FUNCTION_BLOCK CASCADE_CONTROL (* Migrated from IEC 61131-3 ST *)
  (* Standard: 61499-2 *)
  (* Version 1.0, 2026-11-06, st2fb *)
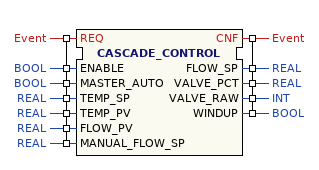
  EVENT_INPUT
    REQ WITH ENABLE, MASTER_AUTO, TEMP_SP, TEMP_PV, FLOW_PV, MANUAL_FLOW_SP;
  END_EVENT
  EVENT_OUTPUT
    CNF WITH FLOW_SP, VALVE_PCT, VALVE_RAW, WINDUP;
  END_EVENT
  VAR_INPUT
    ENABLE : BOOL;
    MASTER_AUTO : BOOL;
    TEMP_SP : REAL;
    TEMP_PV : REAL;
    FLOW_PV : REAL;
    MANUAL_FLOW_SP : REAL;
  END_VAR
  VAR_OUTPUT
    FLOW_SP : REAL;
    VALVE_PCT : REAL;
    VALVE_RAW : INT;
    WINDUP : BOOL;
  END_VAR
  VAR
    M_OUTPUT : REAL;
    M_SAT : BOOL;
    M_RAMP : REAL;
    M_I : REAL;
    M_ERR : REAL;
    M_DEM : REAL;
    S_OUTPUT : REAL;
    S_SAT : BOOL;
    S_RAMP : REAL;
    S_I : REAL;
    S_ERR : REAL;
    S_DEM : REAL;
  END_VAR
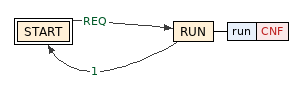
  EC_STATES
    START;
    RUN : run -> CNF;
  END_STATES
  EC_TRANSITIONS
    START TO RUN := REQ;
    RUN TO START := 1;
  END_TRANSITIONS
  ALGORITHM run IN ST:
IF NOT (ENABLE AND MASTER_AUTO) THEN
  M_I := 0.0;
  M_OUTPUT := 0.0;
  M_SAT := FALSE;
ELSE
  IF TEMP_SP > M_RAMP + 2.0 THEN
    M_RAMP := M_RAMP + 2.0;
  ELSIF TEMP_SP < M_RAMP - 2.0 THEN
    M_RAMP := M_RAMP - 2.0;
  ELSE
    M_RAMP := TEMP_SP;
  END_IF;
  M_ERR := M_RAMP - TEMP_PV;
  M_DEM := 0.5 * (1.0 + ABS(M_ERR) ** 0.5) * M_ERR + M_I + 0.125 * M_ERR;
  IF M_DEM > 80.0 THEN
    M_OUTPUT := 80.0;
    M_SAT := TRUE;
  ELSIF M_DEM < 0.0 THEN
    M_OUTPUT := 0.0;
    M_SAT := TRUE;
  ELSE
    M_OUTPUT := M_DEM;
    M_SAT := FALSE;
    M_I := M_I + 0.125 * M_ERR;
  END_IF;
END_IF;
IF MASTER_AUTO THEN
  FLOW_SP := M_OUTPUT;
ELSE
  FLOW_SP := MANUAL_FLOW_SP;
END_IF;
IF NOT ENABLE THEN
  S_I := 0.0;
  S_OUTPUT := 0.0;
  S_SAT := FALSE;
ELSE
  IF FLOW_SP > S_RAMP + 8.0 THEN
    S_RAMP := S_RAMP + 8.0;
  ELSIF FLOW_SP < S_RAMP - 8.0 THEN
    S_RAMP := S_RAMP - 8.0;
  ELSE
    S_RAMP := FLOW_SP;
  END_IF;
  S_ERR := S_RAMP - FLOW_PV;
  S_DEM := 0.25 * (1.0 + ABS(S_ERR) ** 0.5) * S_ERR + S_I + 0.25 * S_ERR;
  IF S_DEM > 100.0 THEN
    S_OUTPUT := 100.0;
    S_SAT := TRUE;
  ELSIF S_DEM < 0.0 THEN
    S_OUTPUT := 0.0;
    S_SAT := TRUE;
  ELSE
    S_OUTPUT := S_DEM;
    S_SAT := FALSE;
    S_I := S_I + 0.25 * S_ERR;
  END_IF;
END_IF;
VALVE_PCT := S_OUTPUT;
VALVE_RAW := REAL_TO_INT(VALVE_PCT * 276.48);
WINDUP := M_SAT OR S_SAT;
  END_ALGORITHM
END_FUNCTION_BLOCK
